// TIA Portal V20 export
// export: Created 2026-10-20T18:54:18.5759495Z, ExportSetting None, DisplayName Totally Integrated Automation Portal, DisplayVersion V20 Update 6, DisplayName TIA Portal Openness, DisplayVersion V20 Update 6, DisplayName TIA Portal Version Control Interface, DisplayVersion V20 Update 6, DisplayName SINAMICS Startdrive Advanced, DisplayVersion V20 SP1, DisplayName SINAMICS Startdrive G130, G150, S120, S150, SINAMICS MV, G220, S200, S210, DisplayVersion V20 SP1, DisplayName SINAMICS Startdrive G110M, G120, G120C, G120D, G120P, G115D, DisplayVersion V20 SP1, DisplayName STEP 7 Professional, DisplayVersion V20 Update 6, DisplayName STEP 7 Safety, DisplayVersion V20 Update 2, DisplayName WinCC Basic/Comfort/Advanced, DisplayVersion V20 Update 6, DisplayName WinCC Unified, DisplayVersion V20 Update 6
VAR_GLOBAL   // PLC tag table "IO_Charger Panels"
   "Charger 1 Contactor ON(1)" AT %I38.0 : Bool;
   "Charger 2 Contactor ON(1)" AT %I38.1 : Bool;
   "Charger 3 Contactor ON(1)" AT %I38.2 : Bool;
   "Charger 1 MCB Helthy(1)" AT %I38.3 : Bool;
   "Charger 2 MCB Helthy(1)" AT %I38.4 : Bool;
   "Charger 3 MCB Helthy(1)" AT %I38.5 : Bool;
   "Charger 1 contactor(1)" AT %Q38.0 : Bool;
   "Charger 2 contactor(1)" AT %Q38.1 : Bool;
   "Charger 3 contactor(1)" AT %Q38.2 : Bool;
   "Charger 1 Contactor ON(2)" AT %I40.0 : Bool;
   "Charger 2 Contactor ON(2)" AT %I40.1 : Bool;
   "Charger 3 Contactor ON(2)" AT %I40.2 : Bool;
   "Charger 1 MCB Helthy(2)" AT %I40.3 : Bool;
   "Charger 2 MCB Helthy(2)" AT %I40.4 : Bool;
   "Charger 3 MCB Helthy(2)" AT %I40.5 : Bool;
   "Charger 1 Contactor ON(3)" AT %I42.0 : Bool;
   "Charger 2 Contactor ON(3)" AT %I42.1 : Bool;
   "Charger 3 Contactor ON(3)" AT %I42.2 : Bool;
   "Charger 1 MCB Helthy(3)" AT %I42.3 : Bool;
   "Charger 2 MCB Helthy(3)" AT %I42.4 : Bool;
   "Charger 3 MCB Helthy(3)" AT %I42.5 : Bool;
   "Charger 1 Contactor ON(4)" AT %I90.0 : Bool;
   "Charger 2 Contactor ON(4)" AT %I90.1 : Bool;
   "Charger 3 Contactor ON(4)" AT %I90.2 : Bool;
   "Charger 1 MCB Helthy(4)" AT %I90.3 : Bool;
   "Charger 2 MCB Helthy(4)" AT %I90.4 : Bool;
   "Charger 3 MCB Helthy(4)" AT %I90.5 : Bool;
   "Charger 1 Contactor ON(5)" AT %I92.0 : Bool;
   "Charger 2 Contactor ON(5)" AT %I92.1 : Bool;
   "Charger 3 Contactor ON(5)" AT %I92.2 : Bool;
   "Charger 1 MCB Helthy(5)" AT %I92.3 : Bool;
   "Charger 2 MCB Helthy(5)" AT %I92.4 : Bool;
   "Charger 3 MCB Helthy(5)" AT %I92.5 : Bool;
   "Charger 1 Contactor ON(6)" AT %I94.0 : Bool;
   "Charger 2 Contactor ON(6)" AT %I94.1 : Bool;
   "Charger 3 Contactor ON(6)" AT %I94.2 : Bool;
   "Charger 1 MCB Helthy(6)" AT %I94.3 : Bool;
   "Charger 2 MCB Helthy(6)" AT %I94.4 : Bool;
   "Charger 3 MCB Helthy(6)" AT %I94.5 : Bool;
   "Charger 1 Contactor ON(7)" AT %I158.0 : Bool;
   "Charger 1 Contactor ON(8)" AT %I160.0 : Bool;
   "Charger 1 contactor(2)" AT %Q39.0 : Bool;
   "Charger 1 contactor(3)" AT %Q196.0 : Bool;
   "Charger 1 contactor(4)" AT %Q197.0 : Bool;
   "Charger 1 contactor(5)" AT %Q236.0 : Bool;
   "Charger 1 contactor(6)" AT %Q301.0 : Bool;
   "Charger 1 contactor(7)" AT %Q367.0 : Bool;
   "Charger 1 contactor(8)" AT %Q368.0 : Bool;
   "Charger 1 MCB Helthy(7)" AT %I158.3 : Bool;
   "Charger 1 MCB Helthy(8)" AT %I160.3 : Bool;
   "Charger 2 Contactor ON(7)" AT %I158.1 : Bool;
   "Charger 2 Contactor ON(8)" AT %I160.1 : Bool;
   "Charger 2 contactor(2)" AT %Q39.1 : Bool;
   "Charger 2 contactor(3)" AT %Q196.1 : Bool;
   "Charger 2 contactor(4)" AT %Q197.1 : Bool;
   "Charger 2 contactor(5)" AT %Q236.1 : Bool;
   "Charger 2 contactor(6)" AT %Q301.1 : Bool;
   "Charger 2 contactor(7)" AT %Q367.1 : Bool;
   "Charger 2 contactor(8)" AT %Q368.1 : Bool;
   "Charger 2 MCB Helthy(7)" AT %I158.4 : Bool;
   "Charger 2 MCB Helthy(8)" AT %I160.4 : Bool;
   "Charger 3 Contactor ON(7)" AT %I158.2 : Bool;
   "Charger 3 Contactor ON(8)" AT %I160.2 : Bool;
   "Charger 3 contactor(2)" AT %Q39.2 : Bool;
   "Charger 3 contactor(3)" AT %Q196.2 : Bool;
   "Charger 3 contactor(4)" AT %Q197.2 : Bool;
   "Charger 3 contactor(5)" AT %Q236.2 : Bool;
   "Charger 3 contactor(6)" AT %Q301.2 : Bool;
   "Charger 3 contactor(7)" AT %Q367.2 : Bool;
   "Charger 3 contactor(8)" AT %Q368.2 : Bool;
   "Charger 3 MCB Helthy(7)" AT %I158.5 : Bool;
   "Charger 3 MCB Helthy(8)" AT %I160.5 : Bool;
END_VAR
